SUBAPPLICATION RedGreenBackground4_AXC (* Hintergrundfarbe (TRUE -> Rot, FALSE -> Grün) für 4 Objekte (AX-Adapter) (Kompakt) *)
  (* Standard: 61499-2 *)
  (* Version 1.0, 2026-07-21, franz, Meisterschulen am Ostbahnhof *)
  PACKAGE MyLib::sys;
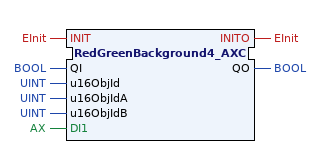
  EVENT_INPUT
    INIT : EInit; (* Initialization Request *)
  END_EVENT
  EVENT_OUTPUT
    INITO : EInit; (* Initialization Confirm *)
  END_EVENT
  VAR_INPUT
    QI : BOOL := TRUE; (* Quality Input - TRUE to enable service *)
    u16ObjId : UINT;
    u16ObjIdA : UINT;
    u16ObjIdB : UINT;
  END_VAR
  VAR_OUTPUT
    QO : BOOL; (* Quality Output - TRUE if service executed successfully *)
  END_VAR
  SOCKETS
    DI1 : adapter::types::unidirectional::AX;
  END_SOCKETS
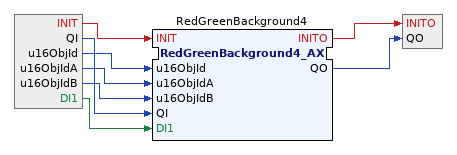
  SUBAPPS
    RedGreenBackground4 : MyLib::sys::RedGreenBackground4_AX;
  END_SUBAPPS
  EVENT_CONNECTIONS
    INIT TO RedGreenBackground4.INIT;
    RedGreenBackground4.INITO TO INITO;
  END_CONNECTIONS
  DATA_CONNECTIONS
    u16ObjId TO RedGreenBackground4.u16ObjId;
    u16ObjIdA TO RedGreenBackground4.u16ObjIdA;
    u16ObjIdB TO RedGreenBackground4.u16ObjIdB;
    QI TO RedGreenBackground4.QI;
    RedGreenBackground4.QO TO QO;
  END_CONNECTIONS
  ADAPTER_CONNECTIONS
    DI1 TO RedGreenBackground4.DI1;
  END_CONNECTIONS
END_SUBAPPLICATION
